Fanuc KAREL source: ka00010.KL

-- PROVISIONAL review KL for V770-1; original PC SHA256 980b4691194ab584ca6d61374f159cd0633be4d379337d1aa7233a8e4be5aae5
-- Incomplete behavior may be omitted. Consult companion uncertainty JSON. Do not deploy.
PROGRAM KA00010
%NOLOCKGROUP
VAR
  SRC : INTEGER
-- UNRESOLVED_DECL DST type=00001c
BEGIN
  -- UNRESOLVED_PC offsets 5-16; opcodes 2E,23
  -- UNRESOLVED_PC offsets 21-33; opcodes 21,23
  -- UNRESOLVED_PC offsets 38-42; opcodes 7F
END KA00010
